(* IEC 61131-3 sources: rusty/compiler/plc_cfc/fixtures/blocks/valid/action_fb, 1 file *)

(* ---- counter.st ---- *)
FUNCTION_BLOCK counter
VAR_INPUT
    in : DINT;
END_VAR
VAR_OUTPUT
    out : DINT;
END_VAR
END_FUNCTION_BLOCK

ACTIONS
    ACTION increment
        out := out + in;
    END_ACTION
END_ACTIONS
